(* IEC 61131-3 sources: Gen-AI/docs/member2_validation/codesys_release_v1.1/C04_missing_dependency, 1 file *)

(* ---- source.st ---- *)
FUNCTION_BLOCK FB_AgentProbeMissingDependency
VAR
 dep : FB_AgentMissingLibraryProbe_6E79B1;
END_VAR
dep();
END_FUNCTION_BLOCK
